(* IEC 61131-3 sources: Caravan/Archiv/12-04-19/Stations/MachineControl/MachineControl/Network/Water_Net, 1 file *)

(* ---- ONE_Water_Net_Table.st ---- *)
#define OBJECTS_CONFIG

FUNCTION GLOBAL TAB ONE_Water_Net
-1$UINT, 0$UINT,
0$UINT, 0$UINT,

2$UDINT,
TO_UDINT(612432597), "FreshWaterTank_Class", 0$UINT, 0$UINT, 1$UINT,
TO_UDINT(4287776992), "InputChange", 0$UINT, 0$UINT, 1$UINT,

_NO_ATTR, TO_UDINT(1967212822), "FRESHWATERTANK_CLASS1",

_NO_ATTR, TO_UDINT(589930375), "INPUTCHANGE1",

//Internal connections
0$UDINT,
0$UDINT,
0$UDINT,
4$UDINT,
TO_UDINT(0), "Water_25", TO_UDINT(1), "Out1",
TO_UDINT(0), "Water_50", TO_UDINT(1), "Out2",
TO_UDINT(0), "Water_75", TO_UDINT(1), "Out3",
TO_UDINT(0), "Water_100", TO_UDINT(1), "Out4",

//Initialization values
0$UDINT,
0$UDINT,

//Symbolic initialization values
0$UDINT,
0$UDINT,

//Initialization of string values
0$UDINT,
0$UDINT,

//Configuration of tasks (RealTime, Cyclic, Background)
0$UDINT,
0$UDINT,

0$UDINT,
2$UDINT,
TO_UDINT(0), (50)$UDINT, 4194303$DINT, 	//FRESHWATERTANK_CLASS1
TO_UDINT(1), (100)$UDINT, 4194303$DINT, 	//INPUTCHANGE1

0$UDINT,
0$UDINT,

//External connections
0$UDINT,
6$UDINT,
TO_UDINT(0), "Start_Check", C_DIR, TO_UDINT(59516340), "TO1611","Output5",
TO_UDINT(0), "WaterPump", C_DIR, TO_UDINT(2870240081), "DI2031","Input5",
TO_UDINT(1), "Input1", C_DIR, TO_UDINT(2870240081), "DI2031","Input1",
TO_UDINT(1), "Input2", C_DIR, TO_UDINT(2870240081), "DI2031","Input2",
TO_UDINT(1), "Input3", C_DIR, TO_UDINT(2870240081), "DI2031","Input3",
TO_UDINT(1), "Input4", C_DIR, TO_UDINT(2870240081), "DI2031","Input4",

//Magic internal connections
0$UDINT,
0$UDINT,

//Configuration of timeslots of tasks (RealTime, Cyclic)
#ifdef __LSLLDR_TIMESLOTS__
0$UDINT,
0$UDINT,

0$UDINT,
0$UDINT,

#endif //__LSLLDR_TIMESLOTS__

//MultiMaster connections
#ifdef __LSLLDR_MULTIMASTER__
0$UDINT,
0$UDINT,
#endif //__LSLLDR_MULTIMASTER__

//Configuration for task ID (RealTime, CyclicTime)
#ifdef __LSLLDR_TASKID__
"\\\\TASKS2  "
0$UDINT,
0$UDINT,

0$UDINT,
2$UDINT,
(0)$UDINT, 	//FRESHWATERTANK_CLASS1
(0)$UDINT, 	//INPUTCHANGE1

0$UDINT,
0$UDINT,

#endif //__LSLLDR_TASKID__

END_FUNCTION
